(* IEC 61131-3 sources: test/Class/SdiasSDCIMaster (part 2) *)

  if StartInInit = 0 then

    // remember that initialization has still to be done
    b_DoTheInit := TRUE;
    // return that initialization is ready so that next step in SdiasManager can begin
    eModuleInitState := READY;

  else

    eModuleInitState := InitTheModule();

  end_if;

END_FUNCTION

FUNCTION VIRTUAL GLOBAL SdiasSDCIMaster::ConnectEvent
  VAR
  	i       : DINT;
    pPort   : ^t_PortInfo;
  END_VAR

  // if we have a seperate read data access => start both read accesses
  if sAccesses.PDOReadDataAccessExtra.pControlByte then
    if sAccesses.CyclicReadInfoAccessOrCombined.pControlByte then
      sAccesses.CyclicReadInfoAccessOrCombined.pControlByte^.EnableDO := TRUE;
    else
      eInitState := _DOHandleInvalid;
      return;
    end_if;

    if sAccesses.PDOReadDataAccessExtra.pControlByte then
      sAccesses.PDOReadDataAccessExtra.pControlByte^.EnableDO := TRUE;
    else
      eInitState := _DOHandleInvalid;
      return;
    end_if;
  else
    if sAccesses.CyclicReadInfoAccessOrCombined.pControlByte then
      // if there are any PDO read data
      if TotalMappingReadSize then
        // remember the pointer to the PDO data and start the combined access
        sAccesses.pPDOReadData := sAccesses.pCyclicReadInfo + sizeof(t_CyclicReadInfo);
      end_if;

      sAccesses.CyclicReadInfoAccessOrCombined.pControlByte^.EnableDO := TRUE;
    else
      eInitState := _DOHandleInvalid;
      return;
    end_if;
  end_if;

  if sAccesses.pPDOWriteData then
    // start the write access
    if sAccesses.PDOWriteDataAccess.pControlByte then
      sAccesses.PDOWriteDataAccess.pControlByte^.EnableDO := TRUE;
    else
      eInitState := _DOHandleInvalid;
      return;
    end_if;
  end_if;

  // set the pointers of the single ports
  pPort := #aPortInfo[0];
  for i := 0 to (SIOL_MAX_PORTS_SUPPORTED-1) do
    // if this port has read data => set the pointer to it
    if pPort^.PdoMapping.ReadDataLength then
      pPort^.pReadData := #LocalReadPDOBuf[0] + pPort^.PdoMapping.ReadDataStartAddress - SIOL_OFFSET_RT_READ_DATA;
    end_if;

    // if this port has write data => set the pointer to it
    if pPort^.PdoMapping.WriteDataLength then
      pPort^.pWriteData := #LocalWritePDOBuf[0] + pPort^.PdoMapping.WriteDataStartAddress - SIOL_OFFSET_RT_WRITE_DATA;
    end_if;

    pPort += sizeof(t_PortInfo);
  end_for;

  //read client value
  StartInInit := StartInInit.Read() <> 0;

  sSdoData.eInitSSW         := t_InitSSW::_InitVariables;

  eInitState := ClassState  := _NotInitialized;

END_FUNCTION

FUNCTION VIRTUAL SdiasSDCIMaster::GetTaskCfg
	VAR_OUTPUT
		TaskCfg 	: BDINT;
	END_VAR

  // we need a call in realtime prescan, realtime postscan and cyclic
  TaskCfg := SDIAS_TASK_MASK_RT_PRE OR SDIAS_TASK_MASK_RT_POST OR SDIAS_TASK_MASK_CY;

END_FUNCTION

FUNCTION VIRTUAL GLOBAL SdiasSDCIMaster::UpdateRt
  VAR
  	i           : USINT;
    pPort       : ^t_PortInfo;
    TempEvent   : t_EventReadData;
  	MyPara      : CmdStruct;
    MyResult    : results;
    PortState   : t_SDCIPortStateBits;
  END_VAR

  // if there is an input pdo => update the pdo input image
  if TotalMappingReadSize then

    PdoProtection.SectionStart();

    _memcpy(ptr1:=#LocalReadPDOBuf[0], ptr2:=sAccesses.pPDOReadData, cntr:=TotalMappingReadSize);

    PdoProtection.SectionStop();
  end_if;

  // save all data local for faster handling and also for using the bits in other methods
  CyclicInfoTotal := sAccesses.pCyclicReadInfo^;

  // things that need to be done with all connected ports / objects
  pPort := #aPortInfo[0];
  for i := 0 to (SIOL_MAX_PORTS_SUPPORTED-1) do
    if pPort^.pThis & (pPort^.ActPortMode <> _Inactive) then
      // if it's a digital input
      if pPort^.pReadData & (pPort^.ActPortMode = _DigitalInput) & pPort^.pInputServer then
        // update the server value
        pPort^.pInputServer^$DINT := pPort^.pReadData^$SINT AND 1;
      end_if;

      // show port state bits
      if pPort^.pPortStateBits then
        PortState := 0; // reset all the higher bits
        PortState.Operating             := to_bool((CyclicInfoTotal.FlagsRdy2OpAndOperating SHR (4 + i)) AND 1);
        PortState.ReadyToOperate        := to_bool((CyclicInfoTotal.FlagsRdy2OpAndOperating SHR      i ) AND 1);
        PortState.InputProcessDataValid := to_bool((CyclicInfoTotal.RtInfoBits              SHR      i ) AND 1);
        PortState.EventAvailable        := to_bool((CyclicInfoTotal.RtInfoBits              SHR (4 + i)) AND 1);
        PortState.OdeState              := to_bool((CyclicInfoTotal.FlagsOdeAndPde          SHR      i ) AND 1);
        PortState.PdeState              := to_bool((CyclicInfoTotal.FlagsOdeAndPde          SHR (4 + i)) AND 1);
        PortState.DuState               := to_bool((CyclicInfoTotal.FlagsDuAndDsUploaded    SHR      i ) AND 1);
        PortState.DsUploaded            := to_bool((CyclicInfoTotal.FlagsDuAndDsUploaded    SHR (4 + i)) AND 1);

        pPort^.pPortStateBits^ := PortState;
      end_if;

      // show fault bits
      if pPort^.pFaultFlags then
        pPort^.pFaultFlags^ := ((CyclicInfoTotal.FaultFlags$UINT SHR (i * 4)) AND 16#F);

        if pPort^.pFaultFlags^ & pPort^.pFaultFlags^ <> pPort^.udOldFaultFlag then

          MyPara.uiCmd    := CMD_SIOL_DEVICE_INFO_UPDATE;
          MyPara.aPara[1] := aPortInfo[i].VendorID;
          MyPara.aPara[2] := aPortInfo[i].DeviceID$DINT;

          // check if a user override is active
          if aPortInfo[i].OverrideMinCycleTime_us then
            MyPara.aPara[3] := aPortInfo[i].OverrideMinCycleTime_us$DINT;
          else
            MyPara.aPara[3] := aPortInfo[i].MinCycleTime_us$DINT;
          end_if;
          MyPara.aPara[4] := aPortInfo[i].ActPortMode$DINT;

          if aPortInfo[i].Required then
            // show required error on SDCI device
            MyPara.aPara[0] := _RequiredError$DINT;

            aPortInfo[i].pThis^.NewInst(#MyPara, #MyResult);

            // crash
            SetRequiredError();
          else
            // show disconnect on class state
            MyPara.aPara[0] := _NoHardware$DINT;

            aPortInfo[i].pThis^.NewInst(#MyPara, #MyResult);
            //there is no sdci hardware at port
            pPort^.PhysicallyAvailable := FALSE;
          end_if;
        end_if;
        //save old state of fault flags
        pPort^.udOldFaultFlag := pPort^.pFaultFlags^;
      end_if;

      // show direct input (always available when there's an object)
      pPort^.pDirectInputServer^$DINT := (CyclicInfoTotal.DigInState SHR i) AND 1;
    end_if;

    pPort += sizeof(t_PortInfo);
  end_for;

  // show voltage bits
  PowerSupply := CyclicInfoTotal.VoltageState$USINT;

  // save the events (if there is an object for the port of the eventsource)
  TempEvent := CyclicInfoTotal.EventData;

  // if it's a valid event
  if TempEvent.EventDatastate.ValidityState then
    if (TempEvent.EventDatastate AND SIOL_EVENT_COUNTER_MASK) <> OldEventCounter then
      // new event => check if we put it into the local buffer or send it to a port object
      if TempEvent.PortNumber = SIOL_MASTER_PORT_NO then
        // add it to the local buffer
        AddEventToBuffer(#TempEvent.EventDetails);
      else
        // check if there is an object
        if (TempEvent.PortNumber < SIOL_MAX_PORTS_SUPPORTED) & aPortInfo[TempEvent.PortNumber].pThis then
          // add it to an object buffer
          MyPara.uiCmd    := CMD_SIOL_DEVICE_ADD_EVENT;

          // pointer to the event details
          MyPara.aPara[0] := (#TempEvent.EventDetails)$DINT;

          aPortInfo[TempEvent.PortNumber].pThis^.NewInst(#MyPara, #MyResult);
        else
          // event dropped, because there is no object for this port or the given portnumber is too high
          EventDropCounter += 1;
        end_if;
      end_if;

      // remember the event counter
      OldEventCounter := TempEvent.EventDatastate AND SIOL_EVENT_COUNTER_MASK;
    end_if;
  end_if;

END_FUNCTION

FUNCTION VIRTUAL GLOBAL SdiasSDCIMaster::UpdateRtPostScan
  VAR
  	i       : DINT;
    pPort   : ^t_PortInfo;
  END_VAR

  if TotalMappingWriteSize then

    PdoProtection.SectionStart();

    _memcpy(ptr1:=sAccesses.pPDOWriteData, ptr2:=#LocalWritePDOBuf[0], cntr:=TotalMappingWriteSize);

    PdoProtection.SectionStop();

    pPort := #aPortInfo[0];
    for i := 0 to (SIOL_MAX_PORTS_SUPPORTED-1) do
      // if it's a digital output
      if pPort^.pWriteData & (pPort^.ActPortMode = _DigitalOutput) & pPort^.pOutputServer then
        // get the current server value
        pPort^.pWriteData^$SINT := to_sint(pPort^.pOutputServer^$DINT AND 1);
      end_if;
      pPort += sizeof(t_PortInfo);
    end_for;
  end_if;

END_FUNCTION

FUNCTION VIRTUAL GLOBAL SdiasSDCIMaster::UpdateCy
  VAR
  	RetcodeIPR : iprStates;
    RetCodeSDCI : t_SDCIRetCode;
  END_VAR

  if b_DoTheInit then

    RetcodeIPR := InitTheModule();

    if RetcodeIPR = ERROR then
#ifdef HWC_LogValue1
      HWC_LogValue1(this, "@0063 (SdiasSDCIMaster::UpdateCy) Failed to initialize module on SDIAS Place 0x{0} via InitModule-Interface", Place);
#endif

      // if it's an required module => error
      if Required then
        SetRequiredError();
      else
        // set init phase over - another try for initialization is NOT done
        b_DoTheInit := FALSE;
      end_if;

      ClassState := _NotInitialized;

    elsif RetcodeIPR = READY then
      // initialization is successful - no more initialization necessary
      b_DoTheInit := FALSE;
      ClassState := _ClassOk;
    else
      // InitTheModule returns BUSY
    end_if;

  else

    if ClassState = _ClassOk then
      sAutoConnectVars.bReConnectStarted := FALSE;

      // if busy with a service data command
      if sSdoData.AsyState = t_SDCIRetCode::SDCI_Busy then
        case sSdoData.AsyCmdType of
        //***************************************************************************************************
          t_AsyCmdType::SingleAsyTransfer:
            case sSdoData.eResponseState of
            //***************************************************************************************************
              t_ReponseState::_PrepareSendData: // start the sending action (done in newinst)

            //***************************************************************************************************
              t_ReponseState::_SendData,
              t_ReponseState::_Wait4SendResponse,
              t_ReponseState::_GotSendResponse,
              t_ReponseState::_ReadData,
              t_ReponseState::_Wait4ReceiveData,
              t_ReponseState::_GotReceiveData:
                if HandleSdoDataTransfer() = ERROR then
                  // set to idle step
                  sSdoData.eResponseState := t_ReponseState::_PrepareSendData;
                end_if;

            //***************************************************************************************************
              t_ReponseState::_GotAllReceiveData:// we enter this step, when we received the answer with the data

                case sSdoData.SdoReadData.ro_RetCode of
                  _FwOk:
                    // ready
                    sSdoData.AsyState := t_SDCIRetCode::SDCI_Ready_Ok;

                  _InvalidChecksum:
                    // error in request CRC detected by firmware
                    sSdoData.AsyState := t_SDCIRetCode::SDCI_MicroCtrl_InvalidChkSum;

                  _FunctionIdNotSupported:
                    // function not supported by firmware
                    sSdoData.AsyState := t_SDCIRetCode::SDCI_MicroCtrl_FunctionIdNotSupported;

                  _InvalidUsageParameter:
                    // invalid usage of parameters detected by firmware
                    sSdoData.AsyState := t_SDCIRetCode::SDCI_MicroCtrl_InvalidParamUsage;

                  _ServiceNotAvailable:
                    // parameter data transfer not possible
                    sSdoData.AsyState := t_SDCIRetCode::SDCI_MicroCtrl_ServiceNotAvailable;

                  _ApplicationError:
                    // error at the SDCI device
                    sSdoData.AsyState := t_SDCIRetCode::SDCI_MicroCtrl_ApplicationError;

                end_case;

                // set to idle step
                sSdoData.eResponseState := t_ReponseState::_PrepareSendData;

                // Handle Asy Callback
                if sSdoData.pCallBackThis & sSdoData.pCallBackFun then
                  HandleSDOCallback();
                else
                  //save received flag of asy data only if it was no callback
                  sSdoData.bSingleAsyTransferReady  := TRUE;
                  sSdoData.udSingleAsyTransferReady := ops.tAbsolute;
                end_if;

                // Unlock SDO Data
                sigclib_atomic_setU32(pValue:=#sSdoData.DataLock, value:= SSDCIM_SDO_UNLOCK);

            //***************************************************************************************************
            end_case;

        //***************************************************************************************************
          t_AsyCmdType::ModeChange,
          t_AsyCmdType::Reconnect,
          t_AsyCmdType::DelayedEnable:
            AsySSW();

        //***************************************************************************************************
        end_case;
      else //if sSdoData.AsyState is not busy

        //if autoconnect is activated it has priority to HandleSDOFifo() -> between each autoconnect are timeslots for other communication (SIOL_MINIMUM_WAIT4RECONNECT_TIME)
        if sAutoConnectVars.bAutoConnectActive = TRUE then
          //check if a new port scan must be started.
          RetCodeSDCI := HandleAutoConnect(sAutoConnectVars.usActPortNbr mod SIOL_MAX_PORTS_SUPPORTED);
          //if reconnect failed because asy communication is busy, wait for asy communication is available
          if RetCodeSDCI <> SDCI_Busy then
            //go to next port
            sAutoConnectVars.usActPortNbr += 1;
          end_if;
        end_if;

        // Check if there are SDOs in the FIFO
        HandleSDOFifo();

      end_if;// if busy with a service data command

      if (b_LogAsyCalls.AsyWarnLogDone      = FALSE) &
         (b_LogAsyCalls.DirectAsyAccessUsed = TRUE)  &
         (b_LogAsyCalls.BufferAsyAccessUsed = TRUE) then

        b_LogAsyCalls.AsyWarnLogDone := TRUE;
        LogError(pMsg:= "@0534 (SdiasSDCIMaster::UpdateCy) WARNING: A combination of buffered and unbuffered asynchronous calls has been detected.");

      end_if;

    end_if; // if ClassState = _ClassOk
  end_if; // if b_DoTheInit

END_FUNCTION

FUNCTION SdiasSDCIMaster::CalcChecksum
	VAR_INPUT
		Mode 	: DINT;
	END_VAR
	VAR_OUTPUT
		Result 	: USINT;
	END_VAR
  VAR
  	i     : UDINT;
    pHelp : ^USINT;
    ForEnd: USINT;
  END_VAR

(*
Checksum calculation:
All of the affected bytes are XOR processed byte by byte. The checksum byte is included with value 0.

The validity of the received telegram can be checked by XOR processing all bytes including the checksum byte. The result must be equal to 0.

*)

  Result := 0;

  // depending on the mode the checksum is calculated over a different memory (and also a different part of it)
  case Mode of
//**********************************************************************************************************************************************************
    0: // read => used to verify received data! the returned value of Result has to be 0 to indicate consistent data
      if sSdoData.SdoReadData.LengthOfData <= SIOL_MAX_SDO_DATA_SIZE then
        if sSdoData.SdoReadData.LengthOfData then
          pHelp   := #sSdoData.SdoReadData.aData[SIOL_MAX_SDO_DATA_SIZE-sSdoData.SdoReadData.LengthOfData];
        else
          pHelp   := (#sSdoData.SdoReadData.ParaIndex)$^USINT;
        end_if;

        ForEnd  := sSdoData.SdoReadData.LengthOfData + sizeof(t_ServiceDataArea.ParaIndex) + sizeof(t_ServiceDataArea.ParaSubIndex) + sizeof(t_ServiceDataArea.PortSelection) + sizeof(t_ServiceDataArea.LengthOfData);

        // calculate over data and access info
        for i := 0 to ForEnd-1 do
          Result := Result XOR pHelp^;
          pHelp  += 1;
        end_for;

        // calculate over msg counter, returncode and checksum (should result in 0 if the data are consistent)
        Result := Result XOR sSdoData.SdoReadData.ro_RetCode$USINT XOR sSdoData.SdoReadData.ro_Checksum XOR sSdoData.SdoReadData.ro_MessageCnt;
      else
        LogError("@04F0 (SdiasSDCIMaster::CalcChecksum) Invalid data length value in SDO response");
      end_if;

//**********************************************************************************************************************************************************
    1: // write => used to fill the checksum field when sending data (therefore the checksum is not included in the calculation)
      if sSdoData.SdoWriteData.LengthOfData <= SIOL_MAX_SDO_DATA_SIZE then
        if sSdoData.SdoWriteData.LengthOfData then
          pHelp   := #sSdoData.SdoWriteData.aData[SIOL_MAX_SDO_DATA_SIZE-sSdoData.SdoWriteData.LengthOfData];
        else
          pHelp   := (#sSdoData.SdoWriteData.ParaIndex)$^USINT;
        end_if;

        ForEnd  := sSdoData.SdoWriteData.LengthOfData + sizeof(t_ServiceDataArea.ParaIndex) + sizeof(t_ServiceDataArea.ParaSubIndex) + sizeof(t_ServiceDataArea.PortSelection) + sizeof(t_ServiceDataArea.LengthOfData) + sizeof(t_ServiceDataArea.wo_ActUsage);

        // calculate over data, access info, usage and msg counter
        for i := 0 to ForEnd-1 do
          Result := Result XOR pHelp^;
          pHelp  += 1;
        end_for;

        Result := Result XOR sSdoData.SdoWriteData.wo_MessageCnt;
      else
        LogError("@04F1 (SdiasSDCIMaster::CalcChecksum) Invalid data length value in SDO request");
      end_if;

//**********************************************************************************************************************************************************
  end_case;

END_FUNCTION

FUNCTION SdiasSDCIMaster::InitializeCyclicSSW
	VAR_INPUT
		pPara 	: ^CmdStruct;
		Usage 	: SdiasSDCIMaster::t_ServiceDataUsage;
	END_VAR
	VAR_OUTPUT
		retcode 	: iprStates;
	END_VAR
  VAR
  	localSDOLock : UDINT;
  END_VAR

  retcode := BUSY;

  // If not busy
  localSDOLock := sigclib_atomic_cmpxchgU32(pValue:=#sSdoData.DataLock, cmpVal := SSDCIM_SDO_UNLOCK, newVal := SSDCIM_SDO_LOCK);
  if localSDOLock = SSDCIM_SDO_UNLOCK then

    // if it's not the master port
    if pPara^.aPara[2]$USINT <> SIOL_MASTER_PORT_NO then
      // take the port from the SDCIPort object
      pPara^.aPara[2] := pPara^.aPara[MAXCMDPARA-1];
    end_if;

    // reset some parts of the readdata structure
    sSdoData.SdoReadData.LengthOfData   := 0;
    sSdoData.SdoReadData.ro_Checksum    := 0;

    retcode := InitializeSdoWriteData(Usage:=Usage, ParaIndex:=pPara^.aPara[0]$UINT, ParaSubIndex:=pPara^.aPara[1]$USINT, PortSelection:=pPara^.aPara[2]$USINT, LengthOfData:=pPara^.aPara[3]$USINT, pData:=pPara^.aPara[4]$pVoid);

    sSdoData.pCallBackThis  := NIL;
    sSdoData.pCallBackFun   := NIL;

    if retcode = ERROR then
      // Unlock SDO Channel
      sigclib_atomic_setU32(pValue:=#sSdoData.DataLock, value:= SSDCIM_SDO_UNLOCK);
      return;
    end_if;

    // we're busy now
    sSdoData.AsyState       := t_SDCIRetCode::SDCI_Busy;
    sSdoData.AsyCmdType     := t_AsyCmdType::SingleAsyTransfer;
    sSdoData.eResponseState := t_ReponseState::_SendData;

  end_if;

END_FUNCTION

FUNCTION SdiasSDCIMaster::GetNextParaFromTable
	VAR_INPUT
		pActPortInfo 	: ^SdiasSDCIMaster::t_PortInfo;
	END_VAR

  // if the next parameter still would be valid
  if pActPortInfo^.ActParaNo+1 < pActPortInfo^.NoOfParameters then
    // set the pointer to the next parameter
    pActPortInfo^.pActPara += sizeof(t_ConfigTablePara) + pActPortInfo^.pActPara^.DataLength;
    pActPortInfo^.ActParaNo += 1;
  else
    // otherwise we're done here
    pActPortInfo^.pActPara := NIL;
  end_if;

END_FUNCTION

FUNCTION SdiasSDCIMaster::FindParaInTable
	VAR_INPUT
		pActPortInfo 	: ^SdiasSDCIMaster::t_PortInfo;
		ParaID 	: UDINT;
		ParaSubID 	: UDINT;
	END_VAR
	VAR_OUTPUT
		pParaInfo 	: ^t_ConfigTablePara;
	END_VAR
  VAR
  	pActPara    : ^t_ConfigTablePara;
    ActParaNo   : UDINT;
  END_VAR

  // Default return value no info available
  pParaInfo := NIL;

  // Start the search at the start of the table
  pActPara  := pActPortInfo^.pFirstPara;
  ActParaNo := 0;

  while ( ( pActPara) &
          ( pActPara^.ParaID <= ParaID) ) do

    // Check if paramter was found
    if ( (pActPara^.ParaID    = ParaID) &
         (pActPara^.ParaSubID = ParaSubID) ) then

      // Return the parameter info
      pParaInfo := pActPara;
      return;

    end_if;

    // Get next parameter
    // Do not use GetNextParaFromTable() because pActPortInfo^.pActPara is manupilated in that method.
    // if the next parameter still would be valid
    if ActParaNo+1 < pActPortInfo^.NoOfParameters then
      // set the pointer to the next parameter
      pActPara += sizeof(t_ConfigTablePara) + pActPara^.DataLength;
      ActParaNo += 1;
    else
      // otherwise we're done here
      pActPara := NIL;
    end_if;

  end_while;

END_FUNCTION

FUNCTION VIRTUAL SdiasSDCIMaster::ReceiveSDOResponse
	VAR_INPUT
		eCommand 	: t_SDIAS_SDO_Cmd;
		hOffset 	: HINT;
		usLength 	: USINT;
		eResult 	: iprStates;
		pResponseBuffer 	: ^USINT;
		ResponseLength 	: USINT;
	END_VAR
	VAR_OUTPUT
		ret_code 	: iprStates;
	END_VAR

  ret_code := SdiasBase::ReceiveSDOResponse(eCommand, hOffset, usLength, eResult, pResponseBuffer, ResponseLength);

  // spi access from baseclass
  if bSDOResponseHandle = TRUE then
    return;
  end_if;

  if eResult = READY then

    case eCommand of
    //*****************************************************************************
      SDIAS_SDO_CMD_MEM_WRITE:
        if sSdoData.eResponseState = _Wait4SendResponse then
          sSdoData.eResponseState := _GotSendResponse;
        else
          LogError("@04F2 (SdiasSDCIMaster::ReceiveSDOResponse) Unexpected SDO response received (object is not waiting for a write memory response)");
        end_if;

    //*****************************************************************************
      SDIAS_SDO_CMD_MEM_READ:
        if sSdoData.eResponseState = _Wait4ReceiveData then
          if ResponseLength & (ResponseLength <= SDIAS_MAX_SDO_READ_LENGTH) then
            if ResponseLength = sSdoData.ActDataSize then
              _memcpy(ptr1:=sSdoData.pActData, ptr2:=pResponseBuffer, cntr:=ResponseLength);
              sSdoData.eResponseState := _GotReceiveData;
            else
              LogError("@04F3 (SdiasSDCIMaster::ReceiveSDOResponse) Received unexpected length of SDO Data");
            end_if;
          else
            LogError("@04F4 (SdiasSDCIMaster::ReceiveSDOResponse) Invalid length in SDO response received");
          end_if;
        else
          LogError("@04F5 (SdiasSDCIMaster::ReceiveSDOResponse) Unexpected SDO response received (object is not waiting for a read memory response)");
        end_if;
    //*****************************************************************************
    end_case;

  else
    case eCommand of
      SDIAS_SDO_CMD_MEM_WRITE:
        LogError("@04F7 (SdiasSDCIMaster::ReceiveSDOResponse) Error at write access!");
      SDIAS_SDO_CMD_MEM_READ:
        LogError("@04F8 (SdiasSDCIMaster::ReceiveSDOResponse) Error at read access!");
    end_case;
  end_if;

END_FUNCTION

FUNCTION SdiasSDCIMaster::InitializeSdoWriteData
	VAR_INPUT
		Usage 	: SdiasSDCIMaster::t_ServiceDataUsage;
		ParaIndex 	: UINT;
		ParaSubIndex 	: USINT;
		PortSelection 	: USINT;
		LengthOfData 	: USINT;
		pData 	: ^void;
		pParaInfo 	: ^t_ConfigTablePara;(* := nil *)
	END_VAR
	VAR_OUTPUT
		retcode 	: iprStates;
	END_VAR

  // initialize variables for the cyclic state machine
  sSdoData.SdoWriteData.ParaIndex     := ParaIndex;
  sSdoData.SdoWriteData.ParaSubIndex  := ParaSubIndex;
  sSdoData.SdoWriteData.PortSelection := PortSelection;
  sSdoData.SdoWriteData.LengthOfData  := LengthOfData;
  if sSdoData.SdoWriteData.LengthOfData then
    if pData then
      if sSdoData.SdoWriteData.LengthOfData <= SIOL_MAX_SDO_DATA_SIZE then

        if pParaInfo = NIL & PortSelection < SIOL_MAX_PORTS_SUPPORTED then
          pParaInfo := FindParaInTable( pActPortInfo  := #aPortInfo[PortSelection]
                                      , ParaID        := ParaIndex
                                      , ParaSubID     := ParaSubIndex);
        end_if;

        if CheckEndianSwapNeeded( pParaInfo     := pParaInfo
                                , PortSelection := PortSelection) then
          EndianSwap( pDst := #sSdoData.SdoWriteData.aData[SIOL_MAX_SDO_DATA_SIZE-sSdoData.SdoWriteData.LengthOfData], pSrc:=pData$^USINT, LengthOfData := sSdoData.SdoWriteData.LengthOfData);
        else
          _memcpy(    ptr1 := #sSdoData.SdoWriteData.aData[SIOL_MAX_SDO_DATA_SIZE-sSdoData.SdoWriteData.LengthOfData], ptr2:=pData,                cntr := sSdoData.SdoWriteData.LengthOfData);
        end_if;

      else
        LogError("@04F9 (SdiasSDCIMaster::InitializeSdoWriteData) Invalid LengthOfData");
        retcode := ERROR;
        return;
      end_if;
    else
      LogError("@04FA (SdiasSDCIMaster::InitializeSdoWriteData) Invalid pointer");
      retcode := ERROR;
      return;
    end_if;
  end_if;

  sSdoData.SdoWriteData.wo_ActUsage   := Usage;
  sSdoData.SdoWriteData.wo_MessageCnt += 1;
  sSdoData.SdoWriteData.wo_Checksum   := CalcChecksum(Mode:=1);

  // set RemainingDataSize, pActData and ActDataSize correctly for the first send package

  // at the initialisation we set the remaining size to the complete package that needs to be transferred
  sSdoData.RemainingDataSize  := sSdoData.SdoWriteData.LengthOfData + sizeof(t_ServiceDataArea) - sizeof(t_ServiceDataArea.aData) - sizeof(t_ServiceDataArea.ro_MessageCnt) - sizeof(t_ServiceDataArea.ro_RetCode) - sizeof(t_ServiceDataArea.ro_Checksum);
  sSdoData.pActData           := #sSdoData.SdoWriteData + SIOL_MAX_SDO_DATA_SIZE - sSdoData.SdoWriteData.LengthOfData;
  if sSdoData.RemainingDataSize > SDIAS_MAX_SDO_WRITE_LENGTH then
    // limit the act size to it's maximum
    sSdoData.ActDataSize := SDIAS_MAX_SDO_WRITE_LENGTH;
  else
    // we only need one package
    sSdoData.ActDataSize := sSdoData.RemainingDataSize;
  end_if;

  retcode := READY;

END_FUNCTION

FUNCTION SdiasSDCIMaster::GetSdoReadData
	VAR_INPUT
		pLength 	: ^USINT;
		pData 	: ^void;
		bDoEndianSwap 	: BOOL;(* := FALSE *)
	END_VAR

  // if pointer to length and data is valid
  if pLength & pData then
    pLength^ := sSdoData.SdoReadData.LengthOfData;

    // if there has been returndata at the SDO transfer
    if sSdoData.SdoReadData.LengthOfData then
      // if the length is valid
      if sSdoData.SdoReadData.LengthOfData <= SIOL_MAX_SDO_DATA_SIZE then

        if bDoEndianSwap = TRUE then
          // Endianswap the returndata to the data pointer
          EndianSwap(pDst := pData$^USINT, pSrc := #sSdoData.SdoReadData.aData[SIOL_MAX_SDO_DATA_SIZE-sSdoData.SdoReadData.LengthOfData], LengthOfData := sSdoData.SdoReadData.LengthOfData);
        else
          // copy the returndata to the data pointer
          _memcpy(   ptr1 := pData,        ptr2 := #sSdoData.SdoReadData.aData[SIOL_MAX_SDO_DATA_SIZE-sSdoData.SdoReadData.LengthOfData],         cntr := sSdoData.SdoReadData.LengthOfData);
        end_if;

      else
        LogError("@04F9 (SdiasSDCIMaster::GetSdoReadData) Invalid LengthOfData");
        pLength^ := 0;
      end_if;
    end_if;
  end_if;

END_FUNCTION

FUNCTION SdiasSDCIMaster::HandleSdoDataTransfer
	VAR_OUTPUT
		retcode 	: iprStates;
	END_VAR

  retcode := READY;

  case sSdoData.eResponseState of
  //***************************************************************************************************
//  t_ReponseState::_PrepareSendData: // preparing the send data is done individually outside of the transfer method

  //***************************************************************************************************
    t_ReponseState::_SendData:
      // send data to the module
      StartWriteSDO(hOffset:=SIOL_OFFSET_SERVICE_DATA_AREA + (sSdoData.pActData$UDINT - (#sSdoData.SdoWriteData.aData)$UDINT)$UINT, usLength:=sSdoData.ActDataSize, pWriteBuffer:=sSdoData.pActData$^USINT, eCommand:=SDIAS_SDO_CMD_MEM_WRITE);
      sSdoData.TimeoutStart   := ops.tAbsolute;
      sSdoData.eResponseState := t_ReponseState::_Wait4SendResponse;

  //***************************************************************************************************
    t_ReponseState::_Wait4SendResponse: // wait for the confirmation of the SDIAS Manager
      // check for a timeout
      if (ops.tAbsolute - sSdoData.TimeoutStart) > SIOL_SDO_TIMEOUT then
        LogError("@04FC (SdiasSDCIMaster::HandleSdoDataTransfer) Timeout at writing SDO command (no response at SDIAS received)");
        sSdoData.AsyErrorCode := t_SDCIRetCode::SDCI_TimeoutInComToMicroCtrl;
        retcode := ERROR;
      end_if;

  //***************************************************************************************************
    t_ReponseState::_GotSendResponse: // we enter this step, when we received the answer
      // here we decide if more packages need to be sent
      sSdoData.RemainingDataSize -= sSdoData.ActDataSize;
      sSdoData.pActData          += sSdoData.ActDataSize;

      // if there is more to send
      if sSdoData.RemainingDataSize then
        // another write access is necessary, prepare the variables
        if sSdoData.RemainingDataSize > SDIAS_MAX_SDO_WRITE_LENGTH then
          // limit the act size to it's maximum
          sSdoData.ActDataSize := SDIAS_MAX_SDO_WRITE_LENGTH;
        else
          // last package
          sSdoData.ActDataSize := sSdoData.RemainingDataSize;
        end_if;

        sSdoData.eResponseState := t_ReponseState::_SendData;
      else
        // finished with writing => go to reading the answer

        sSdoData.ResponseTimeoutStart := ops.tAbsolute;

        // reset the retry counter
        sSdoData.RetryCnt             := 0;

        // at the first reading we try to get as much as we can before checking the real length of the receivedata
        sSdoData.RemainingDataSize := 255; // 255 to signal it is the access to check the real size
        sSdoData.ActDataSize       := SDIAS_MAX_SDO_READ_LENGTH;
        sSdoData.pActData          := #sSdoData.SdoReadData + sizeof(t_ServiceDataArea) - SDIAS_MAX_SDO_READ_LENGTH; // set the pointer to the last block

        sSdoData.eResponseState := t_ReponseState::_ReadData;
      end_if;

  //***************************************************************************************************
    t_ReponseState::_ReadData:// we enter this step to start the read access
      // read data from the module
      StartReadSDO(hOffset:=SIOL_OFFSET_SERVICE_DATA_AREA + (sSdoData.pActData$UDINT - (#sSdoData.SdoReadData.aData)$UDINT)$UINT, usLength:=sSdoData.ActDataSize, eCommand:=SDIAS_SDO_CMD_MEM_READ);
      sSdoData.TimeoutStart   := ops.tAbsolute;
      sSdoData.eResponseState := t_ReponseState::_Wait4ReceiveData;

  //***************************************************************************************************
    t_ReponseState::_Wait4ReceiveData:// we wait for the read data
      // check for a timeout
      if (ops.tAbsolute - sSdoData.TimeoutStart) > SIOL_SDO_TIMEOUT then
        LogError("@04FD (SdiasSDCIMaster::HandleSdoDataTransfer) Timeout at reading SDO response (no response at SDIAS received)");
        sSdoData.AsyErrorCode := t_SDCIRetCode::SDCI_TimeoutInComToMicroCtrl;
        retcode := ERROR;
      end_if;

  //***************************************************************************************************
    t_ReponseState::_GotReceiveData:// we enter this step, when we received the answer with the data
      // here we decide if more packages need to be read

      // check if it's the first access to check the real size
      if sSdoData.RemainingDataSize = 255 then
        // first we check for the mirrored message counter (if the received one is the same, we have an answer from the µC)
        if sSdoData.SdoReadData.ro_MessageCnt = sSdoData.SdoWriteData.wo_MessageCnt then

          // check if we're missing something
          if sSdoData.SdoReadData.LengthOfData > (SDIAS_MAX_SDO_READ_LENGTH - (sizeof(t_ServiceDataArea) - sizeof(t_ServiceDataArea.aData))) then
            sSdoData.RemainingDataSize := sSdoData.SdoReadData.LengthOfData - (SDIAS_MAX_SDO_READ_LENGTH - (sizeof(t_ServiceDataArea) - sizeof(t_ServiceDataArea.aData)));

            // start at the lowest address and work our way up
            sSdoData.pActData -= sSdoData.RemainingDataSize;

            if sSdoData.RemainingDataSize > SDIAS_MAX_SDO_READ_LENGTH then
              // limit the act size to it's maximum
              sSdoData.ActDataSize := SDIAS_MAX_SDO_READ_LENGTH;
            else
              // we only need one package
              sSdoData.ActDataSize := sSdoData.RemainingDataSize;
            end_if;

            sSdoData.eResponseState := t_ReponseState::_ReadData;
          else
            if (CalcChecksum(Mode:=0) = 0) then
              // we got everything already
              sSdoData.eResponseState := t_ReponseState::_GotAllReceiveData;
            else
              if sSdoData.RetryCnt = 0 then
                // try 1 more time, because on simple master (CP101/CP102) it could be that the firmware was writing the message while the OS was reading and therefore we got inconsistent data
                sSdoData.RetryCnt += 1;

                // read everything again
                sSdoData.ResponseTimeoutStart := ops.tAbsolute;

                // at the first reading we try to get as much as we can before checking the real length of the receivedata
                sSdoData.RemainingDataSize := 255; // 255 to signal it is the access to check the real size
                sSdoData.ActDataSize       := SDIAS_MAX_SDO_READ_LENGTH;
                sSdoData.pActData          := #sSdoData.SdoReadData + sizeof(t_ServiceDataArea) - SDIAS_MAX_SDO_READ_LENGTH; // set the pointer to the last block

                sSdoData.eResponseState    := t_ReponseState::_ReadData;
              else
                LogError("@04FE (SdiasSDCIMaster::HandleSdoDataTransfer) Incorrect checksum of response data from firmware detected");
                sSdoData.AsyErrorCode := t_SDCIRetCode::SDCI_InvalidChecksumFromMicroCtrl;
                retcode := ERROR;
              end_if;
            end_if;
          end_if;
        else
          // no answer yet => check timeout and then try again
          if (ops.tAbsolute - sSdoData.ResponseTimeoutStart) > SIOL_SDO_RESPONSE_TIMEOUT then
            LogError("@04FF (SdiasSDCIMaster::HandleSdoDataTransfer) Timeout while waiting for answer of SDCI master firmware");
            sSdoData.AsyErrorCode := t_SDCIRetCode::SDCI_TimeoutInComToMicroCtrl;
            retcode := ERROR;
          else
            // try again

            // at the first reading we try to get as much as we can before checking the real length of the receivedata
            sSdoData.RemainingDataSize := 255; // 255 to signal it is the access to check the real size
            sSdoData.ActDataSize       := SDIAS_MAX_SDO_READ_LENGTH;
            sSdoData.pActData          := #sSdoData.SdoReadData + sizeof(t_ServiceDataArea) - SDIAS_MAX_SDO_READ_LENGTH; // set the pointer to the last block

            sSdoData.eResponseState    := t_ReponseState::_ReadData;
          end_if;
        end_if;
      else
        // here it's not the first access to read data from the module
        sSdoData.RemainingDataSize -= sSdoData.ActDataSize;
        sSdoData.pActData          += sSdoData.ActDataSize;

        // if there is more to read
        if sSdoData.RemainingDataSize then
          // another read access is necessary, prepare the variables
          if sSdoData.RemainingDataSize > SDIAS_MAX_SDO_READ_LENGTH then
            // limit the act size to it's maximum
            sSdoData.ActDataSize := SDIAS_MAX_SDO_READ_LENGTH;
          else
            // last package
            sSdoData.ActDataSize := sSdoData.RemainingDataSize;
          end_if;

          sSdoData.eResponseState := t_ReponseState::_ReadData;
        else
          if (CalcChecksum(Mode:=0) = 0) then
            // finished with reading
            sSdoData.eResponseState := t_ReponseState::_GotAllReceiveData;
          else
            if sSdoData.RetryCnt = 0 then
              // try 1 more time, because on simple master (CP101/CP102) it could be that the firmware was writing the message while the OS was reading and therefore we got inconsistent data
              sSdoData.RetryCnt += 1;

              // read everything again
              sSdoData.ResponseTimeoutStart := ops.tAbsolute;

              // at the first reading we try to get as much as we can before checking the real length of the receivedata
              sSdoData.RemainingDataSize := 255; // 255 to signal it is the access to check the real size
              sSdoData.ActDataSize       := SDIAS_MAX_SDO_READ_LENGTH;
              sSdoData.pActData          := #sSdoData.SdoReadData + sizeof(t_ServiceDataArea) - SDIAS_MAX_SDO_READ_LENGTH; // set the pointer to the last block

              sSdoData.eResponseState    := t_ReponseState::_ReadData;
            else
              LogError("@0501 (SdiasSDCIMaster::HandleSdoDataTransfer) Incorrect checksum of response data from firmware detected");
              sSdoData.AsyErrorCode := t_SDCIRetCode::SDCI_InvalidChecksumFromMicroCtrl;
              retcode := ERROR;
            end_if;
          end_if;
        end_if;
      end_if;

  //***************************************************************************************************
//  t_ReponseState::_GotAllReceiveData:// handling of the receive data is done individually outside of the transfer method

  //***************************************************************************************************
  end_case;

END_FUNCTION

FUNCTION SdiasSDCIMaster::AddEventToBuffer
	VAR_INPUT
		pEventDetails 	: ^SdiasSDCIMaster::t_SDCIEventDetails;
	END_VAR

  PdoProtection.SectionStart();

  // always add the new event to the buffer at the write index
  EventBuffer.aEvents[EventBuffer.EventWrIndex] := pEventDetails^;

  EventBuffer.EventWrIndex += 1;

  if EventBuffer.EventWrIndex = SIOL_EVENT_BUFFER_SIZE then
    EventBuffer.EventWrIndex := 0;
  end_if;

  // if the buffer has already been full
  if NbrOfEventsAvailable = SIOL_EVENT_BUFFER_SIZE then
    // also set the read index to the write index (because that is where the oldest entry is now)
    EventBuffer.EventRdIndex := EventBuffer.EventWrIndex;
  else
    // if not => increase the number of entries
    NbrOfEventsAvailable += 1;
  end_if;

  PdoProtection.SectionStop();

END_FUNCTION

FUNCTION VIRTUAL GLOBAL SdiasSDCIMaster::GetEvent
	VAR_OUTPUT
		OldestEventAvailable 	: SdiasSDCIMaster::t_SDCIEventDetails;
	END_VAR

  PdoProtection.SectionStart();

  // if there are events
  if NbrOfEventsAvailable then
    // get the oldest
    OldestEventAvailable := EventBuffer.aEvents[EventBuffer.EventRdIndex];

    // increment the read pointer of the ring buffer
    EventBuffer.EventRdIndex += 1;
    if EventBuffer.EventRdIndex = SIOL_EVENT_BUFFER_SIZE then
      EventBuffer.EventRdIndex := 0;
    end_if;

    // show that there are less events in the buffer
    NbrOfEventsAvailable -= 1;
  else
    // no event available => set the whole return variable to 0
    _memset(dest:=#OldestEventAvailable, usByte:=0, cntr:=sizeof(OldestEventAvailable));
  end_if;

  PdoProtection.SectionStop();

END_FUNCTION

FUNCTION SdiasSDCIMaster::PrepareParaTabAccess
	VAR_INPUT
		pPortInfo 	: ^SdiasSDCIMaster::t_PortInfo;
	END_VAR
  VAR
  	pHelp     : ^UINT;
    Temp      : UINT;
    pBitHelp  : ^t_BitInfo;
  END_VAR

  // extract PDO info (bit offsets and length of every entry) and set data elements of port info (NoOfParameters & pFirstPara)

  // set pointer on info for process data in
  pHelp := pPortInfo^.pCfgTable + sizeof(t_ConfigTable);

  // number of bit infos for process data in
  Temp := pHelp^;
  pHelp += sizeof(UINT);

  if Temp then
    // allocate memory for the info
    pPortInfo^.pFirstPdIn$pVoid := ToStdLib.Malloc(size:=Temp * sizeof(t_BitInfo));
    pBitHelp := pPortInfo^.pFirstPdIn;

    // if there is a pointer => save the number
    if pBitHelp then
      pPortInfo^.PdInBitInfoNo := Temp;
    end_if;

    while Temp do
      // if we have a memory
      if pBitHelp then
        // store the data there
        pBitHelp^ := pHelp^$t_BitInfo;
        pBitHelp += sizeof(t_BitInfo);
      end_if;

      pHelp += sizeof(t_BitInfo);
      Temp -= 1;
    end_while;
  end_if;

  // number of bit infos for process data out
  Temp := pHelp^;
  pHelp += sizeof(UINT);
  if Temp then
    // allocate memory for the info
    pPortInfo^.pFirstPdOut$pVoid := ToStdLib.Malloc(size:=Temp * sizeof(t_BitInfo));
    pBitHelp := pPortInfo^.pFirstPdOut;

    // if there is a pointer => save the number
    if pBitHelp then
      pPortInfo^.PdOutBitInfoNo := Temp;
    end_if;

    while Temp do
      // if we have a memory
      if pBitHelp then
        // store the data there
        pBitHelp^ := pHelp^$t_BitInfo;
        pBitHelp += sizeof(t_BitInfo);
      end_if;

      pHelp += sizeof(t_BitInfo);
      Temp -= 1;
    end_while;
  end_if;

  // pHelp points to the number of parameters (UDINT)
  pPortInfo^.NoOfParameters := pHelp^$UDINT;
  pHelp += sizeof(UDINT);

  // pHelp points to the first parameter
  pPortInfo^.pFirstPara := pHelp$^t_ConfigTablePara;

END_FUNCTION

FUNCTION VIRTUAL GLOBAL SdiasSDCIMaster::DisconnectEvent
  VAR
  	i           : USINT;
    pPort       : ^t_PortInfo;
  	MyPara      : CmdStruct;
    MyResult    : results;
  END_VAR

  // update own state
  SdiasBase::DisconnectEvent();

  FirmwareVersion     := 0;
  CycleTime           := 0;
  PowerSupply         := 0;

  // reset eventbuffer
  NbrOfEventsAvailable     := 0;
  EventBuffer.EventWrIndex := 0;
  EventBuffer.EventRdIndex := 0;

  // update state to NoHardware
  MyPara.uiCmd        := CMD_SIOL_DEVICE_INFO_UPDATE;
  MyPara.aPara[0]     := _NoHardware$DINT;

  // reset the rest of the module info
  _memset(dest:=#MyPara.aPara[1], usByte:=0, cntr:=4*sizeof(DINT));

  // update state of connected modules
  pPort := #aPortInfo[0];
  for i := 0 to (SIOL_MAX_PORTS_SUPPORTED-1) do
    // if there is an object
    if pPort^.pThis then
      // send the command to reset the device info
      pPort^.pThis^.NewInst(#MyPara, #MyResult);
    end_if;

    pPort += sizeof(t_PortInfo);
  end_for;

  // Unlock is set after InitTheModule completed
  sigclib_atomic_setU32(pValue:=#sSdoData.DataLock, value:= SSDCIM_SDO_LOCK);

  HWKVarSizeFIFO1.Disable();

END_FUNCTION

FUNCTION SdiasSDCIMaster::ExtendPostInitTime
	VAR_INPUT
		AdditionalTime 	: UDINT;
	END_VAR
  VAR
  	MyPara          : CmdStruct;
    MyResult        : results;
  END_VAR

  MyPara.uiCmd    := CMD_EXTEND_POST_INIT_TIME;
  MyPara.aPara[0] := AdditionalTime$DINT;

  SdiasIn.NewInst(#MyPara, #MyResult);

END_FUNCTION

FUNCTION SdiasSDCIMaster::SetRequiredError
  VAR
  	MyPara          : CmdStruct;
    MyResult        : results;
  END_VAR

  // show required error also on SDCI master module
  ClassState := _RequiredError;

  // set required error
  MyPara.uiCmd     := _BUS_IF_SET_REQUIRED_ERROR;

  SdiasIn.NewInst(pPara:=#MyPara, pResult:=#MyResult);
  if MyResult.aData[0]$UDINT then
    LogError("@0502 (SdiasSDCIMaster::SetRequiredError) Failed to set required error to BusInterface");
  end_if;

END_FUNCTION

FUNCTION SdiasSDCIMaster::SelectNextDownloadPara
	VAR_INPUT
		AlsoSearchOtherPorts 	: BOOL;(* := TRUE *)
	END_VAR
	VAR_OUTPUT
		Success 	: BOOL;
	END_VAR

  // in this function we select the next download parameter, if there are no more downloadparameters the pActPara at the current port points to NIL

  Success := TRUE;

  // if we already have a valid pointer => choose the next parameter
  if aPortInfo[sSdoData.ActPortSelection].pActPara then
    GetNextParaFromTable(#aPortInfo[sSdoData.ActPortSelection]);
  end_if;

  if aPortInfo[sSdoData.ActPortSelection].pActPara = NIL then
    // if first parameter or module not available => check for skipping
    if (aPortInfo[sSdoData.ActPortSelection].ActParaNo = 0) | (aPortInfo[sSdoData.ActPortSelection].PhysicallyAvailable = FALSE) then
      // while we're not at the end and there is nothing to download (no sdci port, not physically available or no config parameters) => skip the module
      while (sSdoData.ActPortSelection < SIOL_MAX_PORTS_SUPPORTED) &
            ((aPortInfo[sSdoData.ActPortSelection].CfgPortMode <> _SDCI) | (aPortInfo[sSdoData.ActPortSelection].PhysicallyAvailable = FALSE) |
             (aPortInfo[sSdoData.ActPortSelection].pCfgTable = NIL)      | (aPortInfo[sSdoData.ActPortSelection].NoOfParameters = 0)) do

        if AlsoSearchOtherPorts = FALSE then
          Success := FALSE;
          return;
        end_if;

        sSdoData.ActPortSelection += 1;
      end_while;

      // if we're behind the last possible port => nothing more to initialize
      if sSdoData.ActPortSelection = SIOL_MAX_PORTS_SUPPORTED then
        // tell the caller that we're finished here
        Success := FALSE;
        return;
      end_if;
    end_if;

    // now we are on the first parameter and we have a module that is available => set the pointer to the first parameter
    aPortInfo[sSdoData.ActPortSelection].pActPara := aPortInfo[sSdoData.ActPortSelection].pFirstPara;
  end_if;

  // now skip through the parameters until we find a download parameter or there are no more parameters
  while aPortInfo[sSdoData.ActPortSelection].pActPara &
     (((aPortInfo[sSdoData.ActPortSelection].pActPara^.AccessType <> t_ParaAccessType::rw) &
       (aPortInfo[sSdoData.ActPortSelection].pActPara^.AccessType <> t_ParaAccessType::wo)) |
       (aPortInfo[sSdoData.ActPortSelection].pActPara^.DataLength = 0))
       do

    GetNextParaFromTable(#aPortInfo[sSdoData.ActPortSelection]);

  end_while;

  // now if the pointer is still NIL and we're not yet on the last port => call the method again
  if (aPortInfo[sSdoData.ActPortSelection].pActPara = NIL) then
    // if we're already on the last port => there are no more ports to find download parameters, so we can stop searching
    if sSdoData.ActPortSelection = (SIOL_MAX_PORTS_SUPPORTED-1) then
      Success := FALSE;
    else
      // more ports available => try again with the next port
      if AlsoSearchOtherPorts = FALSE then
        Success := FALSE;
        return;
      end_if;

      sSdoData.ActPortSelection += 1;

      Success := SelectNextDownloadPara();
    end_if;
  end_if;

END_FUNCTION

FUNCTION SdiasSDCIMaster::AsySSW
  VAR
  	TempData            : ARRAY [0..SIOL_MAX_SDO_DATA_SIZE-1] OF USINT;
    TempDataLen         : USINT;
    TempFlags           : t_ControlFlags;
    TempStateFlags      : t_StatusFlags;
  	MyPara              : CmdStruct;
    MyResult            : results;
    TempCycleTime       : UINT;
    i                   : DINT;
  END_VAR

  case sSdoData.eAsySSW of
  //**********************************************************************************************************************************************************
    t_AsySSW::_Idle: // nothing: wait for a command

  //**********************************************************************************************************************************************************
    t_AsySSW::_StartDelayedEnable:
      if DelayedEnablePorts then
        // at the first time we enter here
        if DelayedEnablePorts.FirstTime then
          // reset the port number
          sSdoData.ActPortSelection := 0;
          DelayedEnablePorts.FirstTime := FALSE;
        end_if;

        if DelayedEnablePorts AND 1 then
          // head into the step where the enable takes place
          sSdoData.eAsySSW   := t_AsySSW::_SwitchToNewMode;

          // reset response state machine
          sSdoData.eResponseState := t_ReponseState::_PrepareSendData;
        else
          DelayedEnablePorts := DelayedEnablePorts SHR 1;
          sSdoData.ActPortSelection += 1;
        end_if;
      else
        // we're finished
        sSdoData.eAsySSW  := t_AsySSW::_Finished;
      end_if;

  //**********************************************************************************************************************************************************
    t_AsySSW::_StartReconnect:
      // disable port, enable in scanmode, scan for device, if found => disable again, enable in fixed mode and set operate and pdout valid
      sSdoData.eAsySSW   := t_AsySSW::_RecoDisablePortBe4ScanMode;

      // update state to _NotInitialized
      MyPara.uiCmd        := CMD_SIOL_DEVICE_INFO_UPDATE;
      MyPara.aPara[0]     := _NotInitialized$DINT;

      // reset the rest of the module info
      aPortInfo[sSdoData.ActPortSelection].VendorID := 0;
      aPortInfo[sSdoData.ActPortSelection].DeviceID := 0;
      aPortInfo[sSdoData.ActPortSelection].MinCycleTime_us := 0;

      // vendor ID
      MyPara.aPara[1] := aPortInfo[sSdoData.ActPortSelection].VendorID;

      // device ID
      MyPara.aPara[2] := aPortInfo[sSdoData.ActPortSelection].DeviceID$DINT;

      // minimum cycle time
      if aPortInfo[sSdoData.ActPortSelection].OverrideMinCycleTime_us then
        MyPara.aPara[3] := aPortInfo[sSdoData.ActPortSelection].OverrideMinCycleTime_us$DINT;
      else
        MyPara.aPara[3] := aPortInfo[sSdoData.ActPortSelection].MinCycleTime_us$DINT;
      end_if;

      // actual port mode (still Inactive during initialisation)
      MyPara.aPara[4] := t_SDCIPortMode::_Inactive;

      _memset(dest:=#MyPara.aPara[1], usByte:=0, cntr:=4*sizeof(DINT));

      // send the command to reset the device info
      aPortInfo[sSdoData.ActPortSelection].pThis^.NewInst(#MyPara, #MyResult);

      sSdoData.TargetMode      := aPortInfo[sSdoData.ActPortSelection].StartUpMode;

      // reset response state machine
      sSdoData.eResponseState := t_ReponseState::_PrepareSendData;

  //**********************************************************************************************************************************************************
    t_AsySSW::_StartModeChange:
      // if the port is inactive (mode is inactive and operating is false)
      if (aPortInfo[sSdoData.ActPortSelection].ActPortMode = _Inactive) & ((CyclicInfoTotal.FlagsRdy2OpAndOperating SHR (4+sSdoData.ActPortSelection) AND 1) = FALSE) then
        // directly set new mode
        if sSdoData.TargetMode = _Inactive then
          // if we are already inactive but the user wants to switch again to inactive => start the normal routine (set it inactive again)
          sSdoData.eAsySSW := t_AsySSW::_SetPortInactive;
        else
          // continue setting the new mode
          sSdoData.eAsySSW   := t_AsySSW::_ConfigurePort;
        end_if;
      else
        // first of all we need to deactivate the port
        sSdoData.eAsySSW := t_AsySSW::_SetPortInactive;
      end_if;

      // reset response state machine
      sSdoData.eResponseState := t_ReponseState::_PrepareSendData;

//**********************************************************************************************************************************************************
  	t_AsySSW::_RecoDisablePortBe4ScanMode:
      case sSdoData.eResponseState of
      //***************************************************************************************************
        t_ReponseState::_PrepareSendData: // start the sending action

          // prepare the sdo buffer
          TempData[0]       := E_FNCID_SETPORTCNFPAR; // function ID
          TempData[1]       := sSdoData.ActPortSelection; // port number
          TempData[2]       := t_OpModeStates::E_OPMODE_INACTIVE; // operating mode
          TempData[3]       := t_PortCycle::E_PORTCYCLE_FREERN; // port cycle
          TempData[4]$UINT  := 0; // cycle time
          TempData[6]       :=  aPortInfo[sSdoData.ActPortSelection].PdoMapping.ReadDataLength$USINT; // PDConfig LenIn
          TempData[7]       := (aPortInfo[sSdoData.ActPortSelection].PdoMapping.ReadDataStartAddress - SIOL_OFFSET_RT_READ_DATA)$USINT; // PdConfig PosIn
          TempData[8]       := 0; // PdConfig SrcOffsetIn
          TempData[9]       :=  aPortInfo[sSdoData.ActPortSelection].PdoMapping.WriteDataLength$USINT; // PDConfig LenOut
          TempData[10]      := (aPortInfo[sSdoData.ActPortSelection].PdoMapping.WriteDataStartAddress - SIOL_OFFSET_RT_WRITE_DATA)$USINT; // PdConfig PosOut
          TempData[11]      := 0; // PdConfig SrcOffsetOut
          TempData[12]$UINT := 0; // VendorID
          TempData[14]$UDINT:= 0; // DeviceID
//          _strcpy(dest:=#TempData[18], src:="0000000000000000"); // serial number as string
          _memset(dest:=#TempData[18], usByte:=0, cntr:=16); // serial number as string
          TempData[34]      := 0; // Inspection level
          TempData[35]      := 0; // DS activation state
          TempData[36]      := 0; // DS download enable
          TempData[37]      := 0; // DS upload enable
          TempData[38]      := 16#11; // revision ID (v1.1 should work with both device types, v1.0 doesn't work with v1.1 devices)

          TempDataLen := 39;

          InitializeSdoWriteData(Usage:=_SendFunctionCode, ParaIndex:=0, ParaSubIndex:=0, PortSelection:=SIOL_MASTER_PORT_NO, LengthOfData:=TempDataLen, pData:=#TempData[0]);

          sSdoData.eResponseState := t_ReponseState::_SendData;

      //***************************************************************************************************
        t_ReponseState::_SendData,
        t_ReponseState::_Wait4SendResponse,
        t_ReponseState::_GotSendResponse,
        t_ReponseState::_ReadData,
        t_ReponseState::_Wait4ReceiveData,
        t_ReponseState::_GotReceiveData:
          if HandleSdoDataTransfer() = ERROR then
            sSdoData.eAsySSW := _AsyError;
            return;
          end_if;

      //***************************************************************************************************
        t_ReponseState::_GotAllReceiveData:// we enter this step, when we received the answer with the data

          GetSdoReadData(pLength:=#TempDataLen, pData:=#TempData[0]);
          if TempDataLen = 3 then
            // check response data
            if (TempData[0] = (E_FNCID_SETPORTCNFPAR)$USINT) & // check function ID
               (TempData[1] = sSdoData.ActPortSelection)              // check port number
               then

              if (TempData[2] = 0) then // check status code seperately
                // reset response state machine
                sSdoData.eResponseState := t_ReponseState::_PrepareSendData;

                // finished, continue with next step
                sSdoData.eAsySSW := t_AsySSW::_RecoSwitchToDisableModeBe4ScanMode;
              else
                // error at return code
                LogError("@0503 (SdiasSDCIMaster::AsySSW) Error at status code in answer from µC (_DisablePorts)");
                sSdoData.eAsySSW := _AsyError;
                return;
              end_if;
            else
              // unexpected answer data
              LogError("@0504 (SdiasSDCIMaster::AsySSW) Unexpected data in answer from µC: wrong function ID or port number (_DisablePorts)");
              sSdoData.eAsySSW := _AsyError;
              return;
            end_if;
          else
            // invalid length of answer data
            LogError("@0505 (SdiasSDCIMaster::AsySSW) Invalid data length in answer from µC (_DisablePorts)");
            sSdoData.eAsySSW := _AsyError;
            return;
          end_if;

      //***************************************************************************************************
      end_case;

//**********************************************************************************************************************************************************
  	t_AsySSW::_RecoSwitchToDisableModeBe4ScanMode,
    t_AsySSW::_RecoWait4DisableModeBe4ScanMode:
      case sSdoData.eResponseState of
      //***************************************************************************************************
        t_ReponseState::_PrepareSendData: // start the sending action
          TempFlags := 0;
          if sSdoData.eAsySSW = t_AsySSW::_RecoSwitchToDisableModeBe4ScanMode then
  //          TempFlags.Start2Operate := TRUE; // only makes sense if the port is active in SDCI mode
            TempFlags.OperatingMode := TRUE;
          end_if;

          // prepare the sdo buffer
          TempData[0]       := E_FNCID_CNTSTA; // function ID
          for i:= 0 to SIOL_MAX_PORTS_SUPPORTED-1 do
            // activate the disabled mode for our port
            if i = sSdoData.ActPortSelection then
              TempData[1 + i*sizeof(UINT)]$UINT := TempFlags;
            else
              TempData[1 + i*sizeof(UINT)]$UINT := 0;
            end_if;
          end_for;

          if TotalMappingWriteSize then
            _memset(dest:=#TempData[9], usByte:=0, cntr:=TotalMappingWriteSize);
          end_if;

          TempDataLen := 9 + TotalMappingWriteSize;

          InitializeSdoWriteData(Usage:=_SendFunctionCode, ParaIndex:=0, ParaSubIndex:=0, PortSelection:=SIOL_MASTER_PORT_NO, LengthOfData:=TempDataLen, pData:=#TempData[0]);

          sSdoData.eResponseState := t_ReponseState::_SendData;

      //***************************************************************************************************
        t_ReponseState::_SendData,
        t_ReponseState::_Wait4SendResponse,
        t_ReponseState::_GotSendResponse,
        t_ReponseState::_ReadData,
        t_ReponseState::_Wait4ReceiveData,
        t_ReponseState::_GotReceiveData:
          if HandleSdoDataTransfer() = ERROR then
            sSdoData.eAsySSW := _AsyError;
            return;
          end_if;

      //***************************************************************************************************
        t_ReponseState::_GotAllReceiveData:// we enter this step, when we received the answer with the data

          GetSdoReadData(pLength:=#TempDataLen, pData:=#TempData[0]);
          if TempDataLen = 9 then
            // check response data
            if (TempData[0] = (E_FNCID_CNTSTA)$USINT) then // check function ID
              // reset response state machine
              sSdoData.eResponseState := t_ReponseState::_PrepareSendData;

              // if the operating flag is cleared we can continue
              TempStateFlags := TempData[1 + sSdoData.ActPortSelection*sizeof(t_StatusFlags)]$t_StatusFlags;

              // if any operating bit is still set => go to wait for disabled
              if TempStateFlags.Operating = TRUE then

                // set the time mark the first time we send the command to not wait unnecessary
                if sSdoData.eAsySSW = t_AsySSW::_RecoSwitchToDisableModeBe4ScanMode then
                  Wait4DeviceDisableStartTime := ops.tAbsolute;
                end_if;

                sSdoData.eAsySSW   := t_AsySSW::_RecoWait4DisableModeBe4ScanMode;
              else
                // finished, continue with next step
                sSdoData.eAsySSW   := t_AsySSW::_RecoSetScanMode;
              end_if;
            else
              // unexpected answer data
              LogError("@0506 (SdiasSDCIMaster::AsySSW) Unexpected data in answer from µC: wrong function ID or port number (_SwitchToDisableMode)");
              sSdoData.eAsySSW := _AsyError;
              return;
            end_if;
          else
            // invalid length of answer data
            LogError("@0507 (SdiasSDCIMaster::AsySSW) Invalid data length in answer from µC (_SwitchToDisableMode)");
            sSdoData.eAsySSW := _AsyError;
            return;
          end_if;

      //***************************************************************************************************
      end_case;

//**********************************************************************************************************************************************************
  	t_AsySSW::_RecoSetScanMode:
      // if it's a SDCI port, we must wait the time (according to the specification), because some sensors might need it
      if (aPortInfo[sSdoData.ActPortSelection].CfgPortMode = _SDCI) & ((ops.tAbsolute - Wait4DeviceDisableStartTime) < aPortInfo[sSdoData.ActPortSelection].udModeChangeTime) then
        return;
      end_if;

      case sSdoData.eResponseState of
      //***************************************************************************************************
        t_ReponseState::_PrepareSendData: // start the sending action

          // prepare the sdo buffer
          TempData[0]       := E_FNCID_SETPORTCNFPAR; // function ID
          TempData[1]       := sSdoData.ActPortSelection; // port number
          TempData[2]       := t_OpModeStates::E_OPMODE_SCANMODE; // operating mode
          TempData[3]       := t_PortCycle::E_PORTCYCLE_FREERN; // port cycle
          TempData[4]$UINT  := 0; // cycle time
          TempData[6]       :=  aPortInfo[sSdoData.ActPortSelection].PdoMapping.ReadDataLength$USINT; // PDConfig LenIn
          TempData[7]       := (aPortInfo[sSdoData.ActPortSelection].PdoMapping.ReadDataStartAddress - SIOL_OFFSET_RT_READ_DATA)$USINT; // PdConfig PosIn
          TempData[8]       := 0; // PdConfig SrcOffsetIn
          TempData[9]       :=  aPortInfo[sSdoData.ActPortSelection].PdoMapping.WriteDataLength$USINT; // PDConfig LenOut
          TempData[10]      := (aPortInfo[sSdoData.ActPortSelection].PdoMapping.WriteDataStartAddress - SIOL_OFFSET_RT_WRITE_DATA)$USINT; // PdConfig PosOut
          TempData[11]      := 0; // PdConfig SrcOffsetOut
          TempData[12]$UINT := 0; // VendorID
          TempData[14]$UDINT:= 0; // DeviceID
//          _strcpy(dest:=#TempData[18], src:="0000000000000000"); // serial number as string
          _memset(dest:=#TempData[18], usByte:=0, cntr:=16); // serial number as string
          TempData[34]      := 0; // Inspection level (0 = don't care about vendor or device id)
          TempData[35]      := 0; // DS activation state
          TempData[36]      := 0; // DS download enable
          TempData[37]      := 0; // DS upload enable
          TempData[38]      := 16#11; // revision ID (v1.1 should work with both device types, v1.0 doesn't work with v1.1 devices)

          TempDataLen := 39;

          InitializeSdoWriteData(Usage:=_SendFunctionCode, ParaIndex:=0, ParaSubIndex:=0, PortSelection:=SIOL_MASTER_PORT_NO, LengthOfData:=TempDataLen, pData:=#TempData[0]);

          sSdoData.eResponseState := t_ReponseState::_SendData;

      //***************************************************************************************************
        t_ReponseState::_SendData,
        t_ReponseState::_Wait4SendResponse,
        t_ReponseState::_GotSendResponse,
        t_ReponseState::_ReadData,
        t_ReponseState::_Wait4ReceiveData,
        t_ReponseState::_GotReceiveData:
          if HandleSdoDataTransfer() = ERROR then
            sSdoData.eAsySSW := _AsyError;
            return;
          end_if;

      //***************************************************************************************************
        t_ReponseState::_GotAllReceiveData:// we enter this step, when we received the answer with the data

          GetSdoReadData(pLength:=#TempDataLen, pData:=#TempData[0]);
          if TempDataLen = 3 then
            // check response data
            if (TempData[0] = (E_FNCID_SETPORTCNFPAR)$USINT) & // check function ID
               (TempData[1] = sSdoData.ActPortSelection)              // check port number
               then

              if (TempData[2] = 0) then // check status code seperately
                // reset response state machine
                sSdoData.eResponseState := t_ReponseState::_PrepareSendData;

                // finished, continue with next step
                sSdoData.eAsySSW := t_AsySSW::_RecoSwitchToScanMode;
              else
                // error at return code
                LogError("@0508 (SdiasSDCIMaster::AsySSW) Error at status code in answer from µC (_ConfigurePorts)");
                sSdoData.eAsySSW := _AsyError;
                return;
              end_if;
            else
              // unexpected answer data
              LogError("@0509 (SdiasSDCIMaster::AsySSW) Unexpected data in answer from µC: wrong function ID or port number (_ConfigurePorts)");
              sSdoData.eAsySSW := _AsyError;
              return;
            end_if;
          else
            // invalid length of answer data
            LogError("@050B (SdiasSDCIMaster::AsySSW) Invalid data length in answer from µC  (_ConfigurePorts)");
            sSdoData.eAsySSW := _AsyError;
            return;
          end_if;

      //***************************************************************************************************
      end_case;

//**********************************************************************************************************************************************************
  	t_AsySSW::_RecoSwitchToScanMode,
    t_AsySSW::_RecoWait4ScanMode:
      case sSdoData.eResponseState of
      //***************************************************************************************************
        t_ReponseState::_PrepareSendData: // start the sending action
          TempFlags := 0;
          if sSdoData.eAsySSW = t_AsySSW::_RecoSwitchToScanMode then
            TempFlags.Start2Operate := TRUE;
            TempFlags.OperatingMode := TRUE;
          end_if;

          // prepare the sdo buffer
          TempData[0]       := E_FNCID_CNTSTA; // function ID
          for i:= 0 to SIOL_MAX_PORTS_SUPPORTED-1 do
            if i = sSdoData.ActPortSelection then
              // activate the disabled mode for this port
              TempData[1 + i*sizeof(UINT)]$UINT := TempFlags;
            else
              TempData[1 + i*sizeof(UINT)]$UINT := 0;
            end_if;
          end_for;

          if TotalMappingWriteSize then
            _memset(dest:=#TempData[9], usByte:=0, cntr:=TotalMappingWriteSize);
          end_if;

          TempDataLen := 9 + TotalMappingWriteSize;

          InitializeSdoWriteData(Usage:=_SendFunctionCode, ParaIndex:=0, ParaSubIndex:=0, PortSelection:=SIOL_MASTER_PORT_NO, LengthOfData:=TempDataLen, pData:=#TempData[0]);

          sSdoData.eResponseState := t_ReponseState::_SendData;

      //***************************************************************************************************
        t_ReponseState::_SendData,
        t_ReponseState::_Wait4SendResponse,
        t_ReponseState::_GotSendResponse,
        t_ReponseState::_ReadData,
        t_ReponseState::_Wait4ReceiveData,
        t_ReponseState::_GotReceiveData:
          if HandleSdoDataTransfer() = ERROR then
            sSdoData.eAsySSW := _AsyError;
            return;
          end_if;

      //***************************************************************************************************
        t_ReponseState::_GotAllReceiveData:// we enter this step, when we received the answer with the data

          GetSdoReadData(pLength:=#TempDataLen, pData:=#TempData[0]);
          if TempDataLen = 9 then

            // reset response state machine
            sSdoData.eResponseState := t_ReponseState::_PrepareSendData;

            // check response data
            if (TempData[0] = (E_FNCID_CNTSTA)$USINT) then // check function ID

              // if the operating flag is cleared we can continue
              TempStateFlags := TempData[1 + sSdoData.ActPortSelection*sizeof(t_StatusFlags)]$t_StatusFlags;

              // if the operating bit is not set and there is also no fault => go to wait again
              if (aPortInfo[sSdoData.ActPortSelection].CfgPortMode = _SDCI) & (TempStateFlags.Operating = FALSE) &
                 ((TempStateFlags AND 16#F000) = 0) then // no fault
                sSdoData.eAsySSW   := t_AsySSW::_RecoWait4ScanMode; // wait until fault or operating
              else
                aPortInfo[sSdoData.ActPortSelection].biDeviceInfoSub := SIOL_DEVICEINFO_READSUBINDEXES;
                aPortInfo[sSdoData.ActPortSelection].usActSubIndex   := 2; //first Subindex for read of Device Info data
                // finished, continue with next step
                sSdoData.eAsySSW   := t_AsySSW::_RecoGetDeviceInfos;
              end_if;
            else
              // unexpected answer data
              LogError("@050C (SdiasSDCIMaster::AsySSW) Unexpected data in answer from µC: wrong function ID or port number (_SwitchToNewMode)");
              sSdoData.eAsySSW := _AsyError;
              return;
            end_if;
          else
            // invalid length of answer data
            LogError("@050D (SdiasSDCIMaster::AsySSW) Invalid data length in answer from µC (_SwitchToNewMode)");
            sSdoData.eAsySSW := _AsyError;
            return;
          end_if;

      //***************************************************************************************************
      end_case;

//**********************************************************************************************************************************************************
    t_AsySSW::_RecoGetDeviceInfos:

      case sSdoData.eResponseState of
      //***************************************************************************************************
        t_ReponseState::_PrepareSendData: // start the sending action
          // read direct parameter page 1 (device info)
          InitializeSdoWriteData(Usage:=_ReadParaData, ParaIndex:=0, ParaSubIndex:=aPortInfo[sSdoData.ActPortSelection].usActSubIndex+1, PortSelection:=sSdoData.ActPortSelection, LengthOfData:=0, pData:=NIL);

          sSdoData.eResponseState := t_ReponseState::_SendData;

      //***************************************************************************************************
        t_ReponseState::_SendData,
        t_ReponseState::_Wait4SendResponse,
        t_ReponseState::_GotSendResponse,
        t_ReponseState::_ReadData,
        t_ReponseState::_Wait4ReceiveData,
        t_ReponseState::_GotReceiveData:
          if HandleSdoDataTransfer() = ERROR then
            sSdoData.eAsySSW := _AsyError;
            return;
          end_if;

      //***************************************************************************************************
        t_ReponseState::_GotAllReceiveData:// we enter this step, when we received the answer with the data

          // reset response state machine
          sSdoData.eResponseState := t_ReponseState::_PrepareSendData;
          // initialize next step of ssw -> is changed if more parameters must be read
          sSdoData.eAsySSW := t_AsySSW::_RecoUpdateDeviceObjInfo;

          GetSdoReadData(pLength:=#TempDataLen, pData:=#TempData[0]);
          if (sSdoData.SdoReadData.ro_RetCode = _ServiceNotAvailable) | (TempDataLen = 0) then
            // maybe the port is not connected => select next port (after this if block)
            aPortInfo[sSdoData.ActPortSelection].PhysicallyAvailable := FALSE;

          else
#ifdef SIOL_ENABLE_DEBUG_LOGGING
if TempData$t_DeviceInfoAnswer.ProcessDataIn <> aPortInfo[sSdoData.ActPortSelection].PdoMapping.ReadDataBitLength then
  LogValue("@DBG (SdiasSDCIMaster::AsySSW) Info: Configured bit size of read PDO 0x{0} does not match the expected size from the module 0x{1}. SDCI Port 0x{2}", udValue:=aPortInfo[sSdoData.ActPortSelection].PdoMapping.ReadDataBitLength, udValue2:=TempData$t_DeviceInfoAnswer.ProcessDataIn, udValue3:=sSdoData.ActPortSelection);
end_if;
if TempData$t_DeviceInfoAnswer.ProcessDataOut <> aPortInfo[sSdoData.ActPortSelection].PdoMapping.WriteDataBitLength then
  LogValue("@DBG (SdiasSDCIMaster::AsySSW) Info: Configured bit size of write PDO 0x{0} does not match the expected size from the module 0x{1}. SDCI Port 0x{2}", udValue:=aPortInfo[sSdoData.ActPortSelection].PdoMapping.WriteDataBitLength, udValue2:=TempData$t_DeviceInfoAnswer.ProcessDataOut, udValue3:=sSdoData.ActPortSelection);
end_if;
#endif
            //store act device info read data
            aPortInfo[sSdoData.ActPortSelection].aDeviceInfo[aPortInfo[sSdoData.ActPortSelection].usActSubIndex] := TempData[0];
            //set to next subindex
            aPortInfo[sSdoData.ActPortSelection].usActSubIndex += 1;

            //check for next subindex which must be read
            while aPortInfo[sSdoData.ActPortSelection].usActSubIndex < sizeof(t_DeviceInfoAnswer) do
              if (aPortInfo[sSdoData.ActPortSelection].biDeviceInfoSub shr aPortInfo[sSdoData.ActPortSelection].usActSubIndex) and 0x0001 = TRUE then
                //found next subindex to read
                exit;
              end_if;
              //set entry to next subindex
              aPortInfo[sSdoData.ActPortSelection].usActSubIndex += 1;
            end_while;

            if aPortInfo[sSdoData.ActPortSelection].usActSubIndex < sizeof(t_DeviceInfoAnswer) then
              //read next parameter
              sSdoData.eAsySSW := t_AsySSW::_RecoGetDeviceInfos;
            else
              //finished get device infos
              // MIN CYCLE TIME
              case aPortInfo[sSdoData.ActPortSelection].aDeviceInfo$t_DeviceInfoAnswer.MinCycleTime SHR 6 of
                0: // base of  100µs (Multiplier x time base)
                  aPortInfo[sSdoData.ActPortSelection].MinCycleTime_us :=  100 * (aPortInfo[sSdoData.ActPortSelection].aDeviceInfo$t_DeviceInfoAnswer.MinCycleTime AND 16#3F);

                1: // base of  400µs (Multiplier x time base) +  6400µs
                  aPortInfo[sSdoData.ActPortSelection].MinCycleTime_us :=  400 * (aPortInfo[sSdoData.ActPortSelection].aDeviceInfo$t_DeviceInfoAnswer.MinCycleTime AND 16#3F) +  6400;

                2: // base of 1600µs (Multiplier x time base) + 32000µs
                  aPortInfo[sSdoData.ActPortSelection].MinCycleTime_us := 1600 * (aPortInfo[sSdoData.ActPortSelection].aDeviceInfo$t_DeviceInfoAnswer.MinCycleTime AND 16#3F) + 32000;

                3: // this is reserved for future use
                  LogError("@050E (SdiasSDCIMaster::AsySSW) Invalid time base 3 received at minimum cycle time of device (_GetDeviceInfos)");
                  sSdoData.eAsySSW := _AsyError;
                  return;
              end_case;

              // VENDOR ID
              aPortInfo[sSdoData.ActPortSelection].VendorID := aPortInfo[sSdoData.ActPortSelection].aDeviceInfo$t_DeviceInfoAnswer.VendorIdLsb OR (aPortInfo[sSdoData.ActPortSelection].aDeviceInfo$t_DeviceInfoAnswer.VendorIdMsb SHL 8);

              // DEVICE ID
              aPortInfo[sSdoData.ActPortSelection].DeviceID := aPortInfo[sSdoData.ActPortSelection].aDeviceInfo$t_DeviceInfoAnswer.DeviceIdLsb OR (aPortInfo[sSdoData.ActPortSelection].aDeviceInfo$t_DeviceInfoAnswer.DeviceIdMiddleByte SHL 8) OR (aPortInfo[sSdoData.ActPortSelection].aDeviceInfo$t_DeviceInfoAnswer.DeviceIdMsb SHL 16);

              // Revision ID
              aPortInfo[sSdoData.ActPortSelection].RevisionID := aPortInfo[sSdoData.ActPortSelection].aDeviceInfo$t_DeviceInfoAnswer.RevisionID;

            end_if;
          end_if;

      //***************************************************************************************************
      end_case;

//**********************************************************************************************************************************************************
    t_AsySSW::_RecoUpdateDeviceObjInfo:

      // show the info at the object and also set the class state server

      // reset act parameter number for next init step
      aPortInfo[sSdoData.ActPortSelection].ActParaNo := 0;

      // if there is an object to update
      if aPortInfo[sSdoData.ActPortSelection].pThis then

        // command for the newinst call
        MyPara.uiCmd    := CMD_SIOL_DEVICE_INFO_UPDATE;

        // if it's SDCI device
        if (aPortInfo[sSdoData.ActPortSelection].CfgPortMode = _SDCI) then

          // if there is an IODD file
          if aPortInfo[sSdoData.ActPortSelection].pCfgTable then
            // class state
            if (aPortInfo[sSdoData.ActPortSelection].MinCycleTime_us | aPortInfo[sSdoData.ActPortSelection].OverrideMinCycleTime_us) & aPortInfo[sSdoData.ActPortSelection].VendorID & aPortInfo[sSdoData.ActPortSelection].DeviceID then

              // device available => check if it's the right one
              if (aPortInfo[sSdoData.ActPortSelection].VendorID = aPortInfo[sSdoData.ActPortSelection].pCfgTable^.VendorID) & (aPortInfo[sSdoData.ActPortSelection].DeviceID = aPortInfo[sSdoData.ActPortSelection].pCfgTable^.DeviceID) then
                // show that we are still initializing
                MyPara.aPara[0] := _NotInitialized$DINT;
                aPortInfo[sSdoData.ActPortSelection].PhysicallyAvailable := TRUE;
              else
                // wrong device
                MyPara.aPara[0] := _WrongHardware$DINT;

                // with this it doesn't get enabled when the fixed mode is set on all ports (doesn't make sense if it's the wrong module)
                aPortInfo[sSdoData.ActPortSelection].PhysicallyAvailable := FALSE;
              end_if;
            else
              // device not available
              MyPara.aPara[0] := _NoHardware$DINT;

              aPortInfo[sSdoData.ActPortSelection].PhysicallyAvailable := FALSE;
            end_if;
          else
            // no IODD file => any device is ok if one of the Device Infos is available
            if aPortInfo[sSdoData.ActPortSelection].MinCycleTime_us | aPortInfo[sSdoData.ActPortSelection].OverrideMinCycleTime_us | aPortInfo[sSdoData.ActPortSelection].VendorID | aPortInfo[sSdoData.ActPortSelection].DeviceID then
              // show that we are still initializing
              MyPara.aPara[0] := _NotInitialized$DINT;
              aPortInfo[sSdoData.ActPortSelection].PhysicallyAvailable := TRUE;
            else
              // no device infos available
              MyPara.aPara[0] := _NoHardware$DINT;

              aPortInfo[sSdoData.ActPortSelection].PhysicallyAvailable := FALSE;
            end_if;
          end_if;

          // vendor ID
          MyPara.aPara[1] := aPortInfo[sSdoData.ActPortSelection].VendorID;

          // device ID
          MyPara.aPara[2] := aPortInfo[sSdoData.ActPortSelection].DeviceID$DINT;

          // minimum cycle time
          // check if a user override is active
          if aPortInfo[sSdoData.ActPortSelection].OverrideMinCycleTime_us then
            MyPara.aPara[3] := aPortInfo[sSdoData.ActPortSelection].OverrideMinCycleTime_us$DINT;
          else
            MyPara.aPara[3] := aPortInfo[sSdoData.ActPortSelection].MinCycleTime_us$DINT;
          end_if;

          // actual port mode (still Inactive during initialisation)
          MyPara.aPara[4] := t_SDCIPortMode::_Inactive;

          if aPortInfo[sSdoData.ActPortSelection].Required & (MyPara.aPara[0] <> _NotInitialized$DINT) then
            // show required error on SDCI device
            MyPara.aPara[0] := _RequiredError$DINT;
            aPortInfo[sSdoData.ActPortSelection].pThis^.NewInst(#MyPara, #MyResult);

            SetRequiredError();
          else
            aPortInfo[sSdoData.ActPortSelection].pThis^.NewInst(#MyPara, #MyResult);
          end_if;

        elsif (aPortInfo[sSdoData.ActPortSelection].CfgPortMode = _DigitalInput) | (aPortInfo[sSdoData.ActPortSelection].CfgPortMode = _DigitalOutput) then
          // it's always ok here
          MyPara.aPara[0] := _ClassOk$DINT;
          aPortInfo[sSdoData.ActPortSelection].PhysicallyAvailable := TRUE;

          // we're in the desired mode
          aPortInfo[i].ActPortMode := aPortInfo[i].CfgPortMode;

          // the extra info does not exist here
          MyPara.aPara[1] := 0;
          MyPara.aPara[2] := 0;
          MyPara.aPara[3] := 0;

          // actual port mode is already valid here (no further changes on the setting of this port)
          MyPara.aPara[4] := aPortInfo[sSdoData.ActPortSelection].ActPortMode$DINT;

          aPortInfo[sSdoData.ActPortSelection].pThis^.NewInst(#MyPara, #MyResult);
        end_if;
      else
        // no object available => just like if the module was not physically availabe
        aPortInfo[sSdoData.ActPortSelection].PhysicallyAvailable := FALSE;
      end_if;

      if aPortInfo[sSdoData.ActPortSelection].PhysicallyAvailable = TRUE then
        sSdoData.eAsySSW := t_AsySSW::_RecoCheckDownloadParameters;

        DownloadTimeStart := ops.tAbsolute;

        // if the first pointer is not valid, skip until we find a valid pointer
        if aPortInfo[sSdoData.ActPortSelection].pActPara = NIL then
          if SelectNextDownloadPara(FALSE) = FALSE then
            // no download parameters available

            // go to next step
            sSdoData.eAsySSW := t_AsySSW::_SetPortInactive;

            // reset response state machine
            sSdoData.eResponseState := t_ReponseState::_PrepareSendData;
          end_if;
        end_if;
      else
        // we switch the port to inactive
        sSdoData.TargetMode := _Inactive;

        sSdoData.eAsySSW := t_AsySSW::_SetPortInactive;
      end_if;

//**********************************************************************************************************************************************************
    t_AsySSW::_RecoCheckDownloadParameters:

      case sSdoData.eResponseState of
      //***************************************************************************************************
        t_ReponseState::_PrepareSendData: // start the sending action

          // get the details to write the parameter
          if aPortInfo[sSdoData.ActPortSelection].pActPara then

            if aPortInfo[sSdoData.ActPortSelection].pActPara^.AccessType = t_ParaAccessType::wo then
              // Do not read write only parameters and write the parameter directly
              sSdoData.eAsySSW := t_AsySSW::_RecoDownloadParameters;
            else
              // read the parameter first (to check if it already matches the desired value)
              InitializeSdoWriteData(Usage:=_ReadParaData, ParaIndex:=aPortInfo[sSdoData.ActPortSelection].pActPara^.ParaID$UINT, ParaSubIndex:=aPortInfo[sSdoData.ActPortSelection].pActPara^.ParaSubID$USINT, PortSelection:=sSdoData.ActPortSelection, LengthOfData:=0, pData:=NIL);

              sSdoData.eResponseState := t_ReponseState::_SendData;
            end_if;
          end_if;

      //***************************************************************************************************
        t_ReponseState::_SendData,
        t_ReponseState::_Wait4SendResponse,
        t_ReponseState::_GotSendResponse,
        t_ReponseState::_ReadData,
        t_ReponseState::_Wait4ReceiveData,
        t_ReponseState::_GotReceiveData:
          if HandleSdoDataTransfer() = ERROR then
            sSdoData.eAsySSW := _AsyError;
            return;
          end_if;

      //***************************************************************************************************
        t_ReponseState::_GotAllReceiveData:// we enter this step, when we received the answer with the data

          // extend the post init time by the reaction time of the µC (otherwise we would exceed the timeout of the post init if there are many parameters)
          ExtendPostInitTime(AdditionalTime:=ops.tAbsolute - sSdoData.ResponseTimeoutStart);

          // reset response state machine
          sSdoData.eResponseState := t_ReponseState::_PrepareSendData;

          // check response data
          if (sSdoData.SdoReadData.ro_RetCode = _FwOk) then // check returncode

            // check if the value matches our init value
            GetSdoReadData( pLength       := #TempDataLen
                          , pData         := #TempData[0]
                          , bDoEndianSwap := CheckEndianSwapNeeded( pParaInfo     := aPortInfo[sSdoData.ActPortSelection].pActPara
                                                                  , PortSelection := sSdoData.ActPortSelection) );

            // if it's a string, we add the termination 0 to the uploaded data (for the comparison), because we also have it in the table
            if aPortInfo[sSdoData.ActPortSelection].pActPara^.DataType = _Text then
              TempData[TempDataLen] := 0;
              TempDataLen += 1;
            end_if;

            if (aPortInfo[sSdoData.ActPortSelection].pActPara^.DataLength = TempDataLen) then
              if _memcmp(ptr1:=#TempData[0], ptr2:=aPortInfo[sSdoData.ActPortSelection].pActPara + sizeof(t_ConfigTablePara), cntr:=TempDataLen) = 0 then
                // value match => no download necessary
#ifdef SIOL_ENABLE_DEBUG_LOGGING
LogValue("@DBG (SdiasSDCIMaster::AsySSW) Value and length match already, no download needed. ParameterIndex: {0}, ParameterSubIndex: {1}", udValue:=aPortInfo[sSdoData.ActPortSelection].pActPara^.ParaID, udValue2:=aPortInfo[sSdoData.ActPortSelection].pActPara^.ParaSubID);
#endif
              else

                // it's not the same value => download the parameter
                sSdoData.eAsySSW := t_AsySSW::_RecoDownloadParameters;

#ifdef SIOL_ENABLE_DEBUG_LOGGING
LogValue("@DBG (SdiasSDCIMaster::AsySSW) Value mismatch => download new value. ParameterIndex: {0}, ParameterSubIndex: {1}", udValue:=aPortInfo[sSdoData.ActPortSelection].pActPara^.ParaID, udValue2:=aPortInfo[sSdoData.ActPortSelection].pActPara^.ParaSubID);
#endif

                // skip selecting the next parameter, because we need to send the current parameter in the downloadparameters step
                return;
              end_if;
            else
              // length mismatch

              // if it's a string, we send the new value
              if aPortInfo[sSdoData.ActPortSelection].pActPara^.DataType = _Text then

                // it's not the same value => download the parameter
                sSdoData.eAsySSW := t_AsySSW::_RecoDownloadParameters;

#ifdef SIOL_ENABLE_DEBUG_LOGGING
LogValue("@DBG (SdiasSDCIMaster::AsySSW) Length mismatch at string => download new value. ParameterIndex: {0}, ParameterSubIndex: {1}", udValue:=aPortInfo[sSdoData.ActPortSelection].pActPara^.ParaID, udValue2:=aPortInfo[sSdoData.ActPortSelection].pActPara^.ParaSubID);
#endif

                // skip selecting the next parameter, because we need to send the current parameter in the downloadparameters step
                return;
              else
                LogValue("@050F (SdiasSDCIMaster::AsySSW) Length mismatch (type is not string) => value not downloaded. ParameterIndex: {0}, ParameterSubIndex: {1}", udValue:=aPortInfo[sSdoData.ActPortSelection].pActPara^.ParaID, udValue2:=aPortInfo[sSdoData.ActPortSelection].pActPara^.ParaSubID);
              end_if;
            end_if;

            if SelectNextDownloadPara(FALSE) = FALSE then
              // no more download parameters available

              // go to next step
              sSdoData.eAsySSW := t_AsySSW::_SetPortInactive;
            end_if;
          else
            if (sSdoData.SdoReadData.ro_RetCode = _ApplicationError) then
              // if it's an application error, we also have an error code
              LogValue("@0510 (SdiasSDCIMaster::AsySSW) Error at reading parameter(_CheckDownloadParameters). ParameterIndex: {0}, ParameterSubIndex: {1}, ErrorCode: {2}", udValue:=aPortInfo[sSdoData.ActPortSelection].pActPara^.ParaID, udValue2:=aPortInfo[sSdoData.ActPortSelection].pActPara^.ParaSubID, udValue3:=sSdoData.SdoReadData.aData[230]$HINT);
            else
              LogValue("@0510 (SdiasSDCIMaster::AsySSW) Error at reading parameter(_CheckDownloadParameters). ParameterIndex: {0}, ParameterSubIndex: {1}", udValue:=aPortInfo[sSdoData.ActPortSelection].pActPara^.ParaID, udValue2:=aPortInfo[sSdoData.ActPortSelection].pActPara^.ParaSubID);
            end_if;

            // continue with the next parameter
            if SelectNextDownloadPara(FALSE) = FALSE then
              // no more download parameters available

              // go to next step
              sSdoData.eAsySSW := t_AsySSW::_SetPortInactive;
            end_if;
          end_if;

      //***************************************************************************************************
      end_case;

//**********************************************************************************************************************************************************
    t_AsySSW::_RecoDownloadParameters:

      case sSdoData.eResponseState of
      //***************************************************************************************************
        t_ReponseState::_PrepareSendData: // start the sending action

          // get the details to write the parameter
          if aPortInfo[sSdoData.ActPortSelection].pActPara then

            // prepare everything to send the parameter
            TempDataLen := aPortInfo[sSdoData.ActPortSelection].pActPara^.DataLength;
            _memcpy(ptr1:=#TempData[0], ptr2:=aPortInfo[sSdoData.ActPortSelection].pActPara + sizeof(t_ConfigTablePara), cntr:=TempDataLen);

            InitializeSdoWriteData( Usage         := _WriteParaData
                                  , ParaIndex     := aPortInfo[sSdoData.ActPortSelection].pActPara^.ParaID$UINT
                                  , ParaSubIndex  := aPortInfo[sSdoData.ActPortSelection].pActPara^.ParaSubID$USINT
                                  , PortSelection := sSdoData.ActPortSelection, LengthOfData:=TempDataLen, pData:=#TempData[0]
                                  , pParaInfo     := aPortInfo[sSdoData.ActPortSelection].pActPara);

            sSdoData.eResponseState := t_ReponseState::_SendData;
          else
            sSdoData.eAsySSW := _AsyError;
            LogError("@0511 (SdiasSDCIMaster::AsySSW) Conditions for parameter download not met. No valid parameter pointer!");
            return;
          end_if;

      //***************************************************************************************************
        t_ReponseState::_SendData,
        t_ReponseState::_Wait4SendResponse,
        t_ReponseState::_GotSendResponse,
        t_ReponseState::_ReadData,
        t_ReponseState::_Wait4ReceiveData,
        t_ReponseState::_GotReceiveData:
          if HandleSdoDataTransfer() = ERROR then
            sSdoData.eAsySSW := _AsyError;
            return;
          end_if;

      //***************************************************************************************************
        t_ReponseState::_GotAllReceiveData:// we enter this step, when we received the answer with the data

          // extend the post init time by the reaction time of the µC (otherwise we would exceed the timeout of the post init if there are many parameters)
          ExtendPostInitTime(AdditionalTime:=ops.tAbsolute - sSdoData.ResponseTimeoutStart);

          // in general we go back to check the next parameter (unless there are no more parameters)
          sSdoData.eAsySSW := t_AsySSW::_RecoCheckDownloadParameters;

          // reset response state machine
          sSdoData.eResponseState := t_ReponseState::_PrepareSendData;

          // check response data
          if (sSdoData.SdoReadData.ro_RetCode = _FwOk) then // check returncode

#ifdef SIOL_ENABLE_DEBUG_LOGGING
LogValue("@DBG (SdiasSDCIMaster::AsySSW) Successfully downloaded parameter (_DownloadParameters). ParameterIndex: {0}, ParameterSubIndex: {1}", udValue:=aPortInfo[sSdoData.ActPortSelection].pActPara^.ParaID, udValue2:=aPortInfo[sSdoData.ActPortSelection].pActPara^.ParaSubID);
#endif

          elsif (sSdoData.SdoReadData.ro_RetCode = _ApplicationError) then
            // if it's an application error, we also have an error code
            LogValue("@0512 (SdiasSDCIMaster::AsySSW) Error at writing parameter(_DownloadParameters). ParameterIndex: {0}, ParameterSubIndex: {1}, ErrorCode: {2}", udValue:=aPortInfo[sSdoData.ActPortSelection].pActPara^.ParaID, udValue2:=aPortInfo[sSdoData.ActPortSelection].pActPara^.ParaSubID, udValue3:=sSdoData.SdoReadData.aData[230]$HINT);
          else
            LogValue("@0512 (SdiasSDCIMaster::AsySSW) Error at writing parameter(_DownloadParameters). ParameterIndex: {0}, ParameterSubIndex: {1}", udValue:=aPortInfo[sSdoData.ActPortSelection].pActPara^.ParaID, udValue2:=aPortInfo[sSdoData.ActPortSelection].pActPara^.ParaSubID);
          end_if;

          // select the next parameter
          if SelectNextDownloadPara(FALSE) = FALSE then
            // no more download parameters available

            // go to next step
            sSdoData.eAsySSW := t_AsySSW::_SetPortInactive;

          end_if;

      //***************************************************************************************************
      end_case;

//**********************************************************************************************************************************************************
  	t_AsySSW::_SetPortInactive:
      case sSdoData.eResponseState of
      //***************************************************************************************************
        t_ReponseState::_PrepareSendData: // start the sending action

          // prepare the sdo buffer
          TempData[0]       := E_FNCID_SETPORTCNFPAR; // function ID
          TempData[1]       := sSdoData.ActPortSelection; // port number
          TempData[2]       := t_OpModeStates::E_OPMODE_INACTIVE; // operating mode
          TempData[3]       := t_PortCycle::E_PORTCYCLE_FREERN; // port cycle
          TempData[4]$UINT  := 0; // cycle time
          TempData[6]       :=  aPortInfo[sSdoData.ActPortSelection].PdoMapping.ReadDataLength$USINT; // PDConfig LenIn
          TempData[7]       := (aPortInfo[sSdoData.ActPortSelection].PdoMapping.ReadDataStartAddress - SIOL_OFFSET_RT_READ_DATA)$USINT; // PdConfig PosIn
          TempData[8]       := 0; // PdConfig SrcOffsetIn
          TempData[9]       :=  aPortInfo[sSdoData.ActPortSelection].PdoMapping.WriteDataLength$USINT; // PDConfig LenOut
          TempData[10]      := (aPortInfo[sSdoData.ActPortSelection].PdoMapping.WriteDataStartAddress - SIOL_OFFSET_RT_WRITE_DATA)$USINT; // PdConfig PosOut
          TempData[11]      := 0; // PdConfig SrcOffsetOut
          TempData[12]$UINT := 0; // VendorID
          TempData[14]$UDINT:= 0; // DeviceID
//          _strcpy(dest:=#TempData[18], src:="0000000000000000"); // serial number as string
          _memset(dest:=#TempData[18], usByte:=0, cntr:=16); // serial number as string
          TempData[34]      := 0; // Inspection level
          TempData[35]      := 0; // DS activation state
          TempData[36]      := 0; // DS download enable
          TempData[37]      := 0; // DS upload enable
          TempData[38]      := 16#11; // revision ID (v1.1 should work with both device types, v1.0 doesn't work with v1.1 devices)
